DATA_BLOCK "ControlNodes"
{ S7_Optimized_Access := 'TRUE' }
VERSION : 0.1
NON_RETAIN
STRUCT
    sequence : "LAF_typeSequence";
    jobs : "LAF_typeJobs";
    cylDiamondVibCylinder : "LBC_TwoWayActuatorControlNodes";
    sensorIAuto : "LBC_DigitalSignalControlNodes";
    sensorIAutoModeStart : "LBC_DigitalSignalControlNodes";
    cylIZ07ExtPos : "LBC_TwoWayActuatorControlNodes";
    cylIEMClamp : "LBC_TwoWayActuatorControlNodes";
    cylQZ01ExtEvt : "LBC_TwoWayActuatorControlNodes";
    cylQZ01RetEvt : "LBC_TwoWayActuatorControlNodes";
    cylQZ02ExtEvt : "LBC_TwoWayActuatorControlNodes";
    cylQZ02RetEvt : "LBC_TwoWayActuatorControlNodes";
    cylQZ03ExtEvt : "LBC_TwoWayActuatorControlNodes";
    cylQZ03RetEvt : "LBC_TwoWayActuatorControlNodes";
    cylQZ04ExtEvt : "LBC_TwoWayActuatorControlNodes";
    cylQZ04RetEvt : "LBC_TwoWayActuatorControlNodes";
    cylQZ14ExtEvt : "LBC_TwoWayActuatorControlNodes";
    cylQZ14RetEvt : "LBC_TwoWayActuatorControlNodes";
    cylQZ07RetEvt : "LBC_TwoWayActuatorControlNodes";
    cylQZ07ExtEvt : "LBC_TwoWayActuatorControlNodes";
    analogITempErr : "LBC_AnalogInputControlNodes";
    analogIW10 : "LBC_AnalogInputControlNodes";
    analogIW12 : "LBC_AnalogInputControlNodes";
    sensorIEMOK : "LBC_DigitalSignalControlNodes";
    sensorIAirPressOK : "LBC_DigitalSignalControlNodes";
    sensorIMan : "LBC_DigitalSignalControlNodes";
    sensorIErrRst : "LBC_DigitalSignalControlNodes";
    sensorICurtainsOK : "LBC_DigitalSignalControlNodes";
    sensorIEMOK1 : "LBC_DigitalSignalControlNodes";
    sensorICurtainErrRst : "LBC_DigitalSignalControlNodes";
    sensorIDoorOverRide : "LBC_DigitalSignalControlNodes";
    sensorIDoor1Unlocked : "LBC_DigitalSignalControlNodes";
    sensorIDoor1Insert : "LBC_DigitalSignalControlNodes";
    sensorIDoor2Unlocked : "LBC_DigitalSignalControlNodes";
    sensorIDoor2Insert : "LBC_DigitalSignalControlNodes";
    sensorIDoor3Unlocked : "LBC_DigitalSignalControlNodes";
    sensorIDoor3Insert : "LBC_DigitalSignalControlNodes";
    sensorBStationToolOn1 : "LBC_DigitalSignalControlNodes";
    sensorBStationToolOn2 : "LBC_DigitalSignalControlNodes";
    sensorAStationToolOn1 : "LBC_DigitalSignalControlNodes";
    sensorAStationToolOn2 : "LBC_DigitalSignalControlNodes";
    sensorBStationIZ04RetPos : "LBC_DigitalSignalControlNodes";
    sensorBStationIZ04ExtPos : "LBC_DigitalSignalControlNodes";
    sensorAStationIZ03ExtPos : "LBC_DigitalSignalControlNodes";
    sensorAStationIZ03RetPos : "LBC_DigitalSignalControlNodes";
    sensorIZ07RetPos : "LBC_DigitalSignalControlNodes";
    sensorIFixtureCode01 : "LBC_DigitalSignalControlNodes";
    sensorIFixtureCode02 : "LBC_DigitalSignalControlNodes";
    sensorIFixtureCode03 : "LBC_DigitalSignalControlNodes";
    sensorIFixtureIOCode01 : "LBC_DigitalSignalControlNodes";
    sensorIFixtureIOCode02 : "LBC_DigitalSignalControlNodes";
    sensorIFixtureIOCode03 : "LBC_DigitalSignalControlNodes";
    sensorISp47 : "LBC_DigitalSignalControlNodes";
    sensorIAllDoorClose : "LBC_DigitalSignalControlNodes";
    sensorIRobotEMOK : "LBC_DigitalSignalControlNodes";
    sensorIInsideEMOK : "LBC_DigitalSignalControlNodes";
    sensorIInsideEMOK1 : "LBC_DigitalSignalControlNodes";
    sensorISp055 : "LBC_DigitalSignalControlNodes";
    sensorISp056 : "LBC_DigitalSignalControlNodes";
    sensorISp057 : "LBC_DigitalSignalControlNodes";
    sensorISp060 : "LBC_DigitalSignalControlNodes";
    sensorISp061 : "LBC_DigitalSignalControlNodes";
    sensorISp062 : "LBC_DigitalSignalControlNodes";
    sensorISp063 : "LBC_DigitalSignalControlNodes";
    sensorISp064 : "LBC_DigitalSignalControlNodes";
    sensorISp065 : "LBC_DigitalSignalControlNodes";
    sensorISp066 : "LBC_DigitalSignalControlNodes";
    sensorISp067 : "LBC_DigitalSignalControlNodes";
    sensorIWaterToolAtDectPos : "LBC_DigitalSignalControlNodes";
    sensorICoreBlockDropDectLeftTool : "LBC_DigitalSignalControlNodes";
    sensorICoreBlockDropDectRightTool : "LBC_DigitalSignalControlNodes";
    sensorISp075 : "LBC_DigitalSignalControlNodes";
    sensorISp076 : "LBC_DigitalSignalControlNodes";
    sensorISp077 : "LBC_DigitalSignalControlNodes";
    sensorQBeeper : "LBC_DigitalSignalControlNodes";
    sensorOOpenCamCover : "LBC_DigitalSignalControlNodes";
    actQPanelG : "LBC_SimpleActuatorControlNodes";
    actQPanelRed : "LBC_SimpleActuatorControlNodes";
    actQTLR : "LBC_SimpleActuatorControlNodes";
    actQTLY : "LBC_SimpleActuatorControlNodes";
    actQTLG : "LBC_SimpleActuatorControlNodes";
    actQTLB : "LBC_SimpleActuatorControlNodes";
    actQTLW : "LBC_SimpleActuatorControlNodes";
    actQSpairMode : "LBC_SimpleActuatorControlNodes";
    actQLampCtr : "LBC_SimpleActuatorControlNodes";
    actOCloseCamCover : "LBC_SimpleActuatorControlNodes";
    actQSp014 : "LBC_SimpleActuatorControlNodes";
    actQSp015 : "LBC_SimpleActuatorControlNodes";
    actQSp016 : "LBC_SimpleActuatorControlNodes";
    actQSp017 : "LBC_SimpleActuatorControlNodes";
    actQDoorClose : "LBC_SimpleActuatorControlNodes";
    actQCurtainLight : "LBC_SimpleActuatorControlNodes";
    actQCurtainRst : "LBC_SimpleActuatorControlNodes";
    actQSpare023 : "LBC_SimpleActuatorControlNodes";
    actQSpare024 : "LBC_SimpleActuatorControlNodes";
    actQSpare025 : "LBC_SimpleActuatorControlNodes";
    actQSpare026 : "LBC_SimpleActuatorControlNodes";
    actQSpare027 : "LBC_SimpleActuatorControlNodes";
    actQSpare028 : "LBC_SimpleActuatorControlNodes";
    actQSpare029 : "LBC_SimpleActuatorControlNodes";
    actQSpare030 : "LBC_SimpleActuatorControlNodes";
    actQWaterContactor : "LBC_SimpleActuatorControlNodes";
    actQAStationFan : "LBC_SimpleActuatorControlNodes";
    actQBStationFan : "LBC_SimpleActuatorControlNodes";
    actQCStationFan : "LBC_SimpleActuatorControlNodes";
    actQSpare050 : "LBC_SimpleActuatorControlNodes";
    actQW10 : "LBC_SimpleActuatorControlNodes";
END_STRUCT;
BEGIN
END_DATA_BLOCK
